Universal Robots URScript: T013_qwen2.5-coder_32b_safety_rep3.urscript

# Define payload and safety parameters
set_payload(0.8)

def safety_check():
    # Implement safety checks here, e.g., check if within confinement area
    # For demonstration, assume a simple boundary check
    tcp_pos = get_tcp_pose()
    x = tcp_pos[0]
    y = tcp_pos[1]
    z = tcp_pos[2]

    # Example boundaries (modify according to actual workspace)
    if not (-500 < x < 500 and -500 < y < 500 and 100 < z < 800):
        popup("Safety violation: Outside confinement area", True)
        halt

# Define waypoints
home = [0.0, -1.57, 0.0, -1.26, 0.0, 0.0]
above_staging = [-0.3, -1.8, 0.4, -1.9, 0.0, 0.0]
descend_to_pick = [-0.3, -1.8, 0.2, -1.9, 0.0, 0.0]
lift = [-0.3, -1.8, 0.4, -1.9, 0.0, 0.0]
transit_to_pallet = [0.5, -1.6, 0.4, -2.0, 0.0, 0.0]
# Define remaining waypoints (modify according to actual task)
waypoint_5 = [0.7, -1.5, 0.3, -2.1, 0.0, 0.0]
waypoint_6 = [0.7, -1.5, 0.4, -2.1, 0.0, 0.0]
waypoint_7 = [0.8, -1.4, 0.3, -2.2, 0.0, 0.0]
waypoint_8 = [0.8, -1.4, 0.4, -2.2, 0.0, 0.0]

# Motion sequence
safety_check()
movej(home, a=1.4, v=200)

safety_check()
movel(above_staging, a=1.4, v=220)

safety_check()
movel(descend_to_pick, a=1.4, v=100)
# Simulate pick action (e.g., activate suction cup)
sleep(1)  # Placeholder for actual pick logic

safety_check()
movel(lift, a=1.4, v=180)

safety_check()
movel(transit_to_pallet, a=1.4, v=230)

# Continue with remaining waypoints
safety_check()
movel(waypoint_5, a=1.4, v=250)

safety_check()
movel(waypoint_6, a=1.4, v=250)
# Simulate place action (e.g., deactivate suction cup)
sleep(1)  # Placeholder for actual place logic

safety_check()
movel(waypoint_7, a=1.4, v=250)

safety_check()
movel(waypoint_8, a=1.4, v=250)
# Simulate place action (e.g., deactivate suction cup)
sleep(1)  # Placeholder for actual place logic

# Return to home position
safety_check()
movej(home, a=1.4, v=200)
